Staubli VAL3: updateTool.pgx

public program updateTool(num x_nToolNumber, bool x_bOffsetActive)
  local bool l_bOut
  local num l_nStep
begin
  l_bOut=false
  l_nStep=0
  do
    switch l_nStep
      case 0
        //Decide which tool to use
        utCurrentTool.nItem=x_nToolNumber
        switch x_nToolNumber
          case 0
            utCurrentTool.tValue=tFlange
            utLbl_Tool_Data.Common.sText="tFlange"
            //call hmiAlert("SwitchFlange")
            l_nStep=1
          break
          case 1
            utCurrentTool.tValue=tTool1
            utLbl_Tool_Data.Common.sText="tTool1"
            //call hmiAlert("SwitchTool1")
            l_nStep=1
          break
          case 2
            utCurrentTool.tValue=tTool2
            utLbl_Tool_Data.Common.sText="tTool2"
            //call hmiAlert("SwitchTool2")
            l_nStep=1
          break
          case 3
            utCurrentTool.tValue=tTool3
            utLbl_Tool_Data.Common.sText="tTool3"
            //call hmiAlert("SwitchTool3")
            l_nStep=1
          break
        endSwitch
      break
      //
      case 1
        //Add or not add tool deviations?
        if utImg_Switch.Data.bStatus==true and x_bOffsetActive==true
          utCurrentTool.tValue.trsf=utCurrentTool.tValue.trsf*trOffset
          l_nStep=2
        else
          utCurrentTool.tValue.trsf=utCurrentTool.tValue.trsf
          l_nStep=2
        endIf
      break
      //
      case 2
        //Update current tool value
        tCurrentTool=utCurrentTool.tValue
        $jogContext(tCurrentTool,world,0)
        l_nStep=3
      break
      //
      case 3
        l_bOut=true
      break
    endSwitch
  until l_bOut
end
